// TIA Portal V20 export
DATA_BLOCK "02_Wartungszaehler_DB"   // DB4
AUTHOR : Falter
FAMILY : HMI
VERSION : 1.0
// stored: InstanceOfName 02_Wartungszaehler, InstanceOfType FB
"02_Wartungszaehler"
   // VAR
   //    Wartungszähler_Positionierachse_Zyklen : "FB_Wartungszähler_Zyklen";
   //    Wartungszähler_Drehachse_Zyklen : "FB_Wartungszähler_Zyklen";
   //    Wartungszähler_Positionierachse_Weg : "FB_Wartungszähler_Weg";
   //    Wartungszähler_Drehachse_Weg : "FB_Wartungszähler_Weg";
   // END_VAR
   // VAR RETAIN
   //    Positionierachse_Weg { S7_SetPoint := 'True'} : DInt;
   //    Drehachse_Weg { S7_SetPoint := 'True'} : DInt;
   // END_VAR
BEGIN
END_DATA_BLOCK
